Universal Robots URScript: T009_zai-org_GLM-4.7-FP8_edit_perf_rep1.urscript

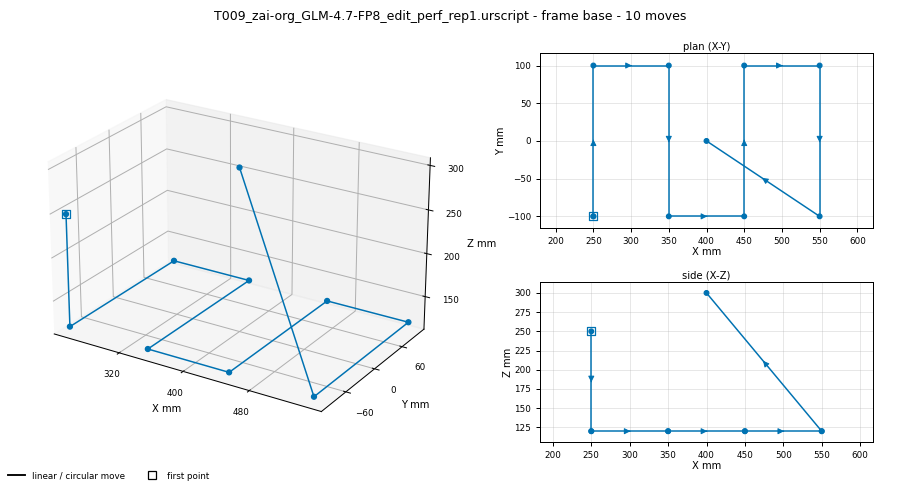
[picture p0: tool path of T009_zai-org_GLM-4.7-FP8_edit_perf_rep1.urscript in frame base, 10 of 12 moves have a stored position in this frame; points joined in program order, loops and branches not executed]
# Task: T009 — Laser surface scan — fenced mode (Optimized)
# Generated by ENFIELD IR→URScript Translator
# Operating mode: fenced | Max TCP speed: 0.200 m/s
# Robot: ur5e
#
# WARNING: This is auto-generated code for SIMULATION ONLY.
# Do NOT deploy to a physical robot without safety review.

def task_T009():
  # [0] Verify E-Stop
  # E-Stop safety check (hardware-enforced on UR controller)
  if (get_digital_in(0) == True):
    popup("E-Stop active — aborting program.", error=True)
    halt
  end

  # [1] Home (Optimized joint speed/accel)
  movej([0.0000, -1.5708, 1.5708, -1.5708, -1.5708, 0.0000], a=2.0000, v=2.0000)

  # [2] Above scan start (Max TCP speed, increased accel, larger blend)
  movel(p[0.250000, -0.100000, 0.250000, 0.0000, 3.1416, 0.0000], a=1.2000, v=0.2000, r=0.0200)

  # [3] Descend to scan height (Max TCP speed, increased accel, larger blend)
  movel(p[0.250000, -0.100000, 0.120000, 0.0000, 3.1416, 0.0000], a=1.2000, v=0.2000, r=0.0200)

  # [4] Laser ON
  set_digital_out(3, True)

  # [5] Scan line 1 (Max TCP speed, increased accel, larger blend)
  movel(p[0.250000, 0.100000, 0.120000, 0.0000, 3.1416, 0.0000], a=1.2000, v=0.2000, r=0.0200)

  # [6] Step to line 2 (Max TCP speed, increased accel, larger blend)
  movel(p[0.350000, 0.100000, 0.120000, 0.0000, 3.1416, 0.0000], a=1.2000, v=0.2000, r=0.0200)

  # [7] Scan line 2 reverse (Max TCP speed, increased accel, larger blend)
  movel(p[0.350000, -0.100000, 0.120000, 0.0000, 3.1416, 0.0000], a=1.2000, v=0.2000, r=0.0200)

  # [8] Step to line 3 (Max TCP speed, increased accel, larger blend)
  movel(p[0.450000, -0.100000, 0.120000, 0.0000, 3.1416, 0.0000], a=1.2000, v=0.2000, r=0.0200)

  # [9] Scan line 3 (Max TCP speed, increased accel, larger blend)
  movel(p[0.450000, 0.100000, 0.120000, 0.0000, 3.1416, 0.0000], a=1.2000, v=0.2000, r=0.0200)

  # [10] Step to line 4 (Max TCP speed, increased accel, larger blend)
  movel(p[0.550000, 0.100000, 0.120000, 0.0000, 3.1416, 0.0000], a=1.2000, v=0.2000, r=0.0200)

  # [11] Scan line 4 reverse (Max TCP speed, increased accel, stop at end)
  movel(p[0.550000, -0.100000, 0.120000, 0.0000, 3.1416, 0.0000], a=1.2000, v=0.2000)

  # [12] Laser OFF
  set_digital_out(3, False)

  # [13] Retract (Max TCP speed, increased accel)
  movel(p[0.400000, 0.000000, 0.300000, 0.0000, 3.1416, 0.0000], a=1.2000, v=0.2000, r=0.0200)

  # [14] Return home (Optimized joint speed/accel)
  movej([0.0000, -1.5708, 1.5708, -1.5708, -1.5708, 0.0000], a=2.0000, v=2.0000)

end

# Entry point
task_T009()
